Yaskawa INFORM job: TURNPRO.JBI

/JOB
//NAME TURNPRO
//POS
///NPOS 9,0,0,0,0,0
///TOOL 9
///POSTYPE PULSE
///PULSE
C00000=360640,0,0,0,27307,0
C00001=0,0,0,-213423,27307,0
C00002=0,0,0,0,27307,112537
C00003=-360640,0,0,0,27307,-112537
C00004=0,369664,-239810,0,172942,0
C00005=-162288,-58368,75729,192081,-27307,-101283
C00006=631120,0,0,-373491,27307,303849
C00007=-324576,0,0,192081,0,-303849
C00008=631120,0,0,-373491,27307,303849
//INST
<volatile>
///COMM Generated using RoboDK
///ATTR SC,RW
///GROUP1 RB1
NOP
'Program generated by RoboDK v
'6.0.7 for Yaskawa Motoman DX1
'350D on XX/XX/XXXX 18:00:00
'Using nominal kinematics.
'Using Frame S (targets wrt ba
'se):
'1234.6,-98.8,50.5,0.0,0.0,30.
'0
'Tool Tool S should be close t
'o:
'10.0,20.0,150.0,0.0,0.0,0.0
MOVL C00000 V=100.0
MOVL C00001 V=100.0
MOVL C00002 V=100.0
MOVL C00003 V=100.0
MOVL C00004 V=100.0
MOVL C00005 V=100.0
MOVL C00006 V=100.0
MOVL C00007 V=100.0
MOVJ C00008 VJ=50.00
END
